FUNCTION FC 1 : VOID
VAR_TEMP
  x : INT;
END_VAR
BEGIN
END_FUNCTION
